(* IEC 61131-3 sources: plc-vscode/tests/st/test-ready/trust-platform/examples/OSCAT/warehouse_conveyor_merge_mediator/oop/src, 3 files *)

(* ---- Main.st ---- *)
(* Pattern role: IInfeedConveyor is the contract boundary for the Mediator example. *)
INTERFACE IInfeedConveyor
    PROPERTY LaneId : INT
    GET
    END_GET
    END_PROPERTY
    PROPERTY Requesting : BOOL
    GET
    END_GET
    END_PROPERTY
    PROPERTY Jammed : BOOL
    GET
    END_GET
    END_PROPERTY
    PROPERTY Granted : BOOL
    GET
    END_GET
    END_PROPERTY
    METHOD UpdateLane
    VAR_INPUT
        Request : BOOL;
        Jam : BOOL;
    END_VAR
    END_METHOD
    METHOD Grant
    VAR_INPUT
        Enable : BOOL;
    END_VAR
    END_METHOD
END_INTERFACE

(* Pattern role: InfeedConveyor is a concrete implementation in the Mediator example. *)
FUNCTION_BLOCK InfeedConveyor IMPLEMENTS IInfeedConveyor
VAR
    LaneIdValue : INT;
    RequestingValue : BOOL;
    JammedValue : BOOL;
    GrantedValue : BOOL;
END_VAR
METHOD PUBLIC Configure
VAR_INPUT
    LaneId : INT;
END_VAR
LaneIdValue := LaneId;
END_METHOD
METHOD PUBLIC UpdateLane
VAR_INPUT
    Request : BOOL;
    Jam : BOOL;
END_VAR
RequestingValue := Request;
JammedValue := Jam;
END_METHOD
METHOD PUBLIC Grant
VAR_INPUT
    Enable : BOOL;
END_VAR
GrantedValue := Enable;
END_METHOD
PUBLIC PROPERTY LaneId : INT
GET
    LaneId := LaneIdValue;
END_GET
END_PROPERTY
PUBLIC PROPERTY Requesting : BOOL
GET
    Requesting := RequestingValue;
END_GET
END_PROPERTY
PUBLIC PROPERTY Jammed : BOOL
GET
    Jammed := JammedValue;
END_GET
END_PROPERTY
PUBLIC PROPERTY Granted : BOOL
GET
    Granted := GrantedValue;
END_GET
END_PROPERTY
END_FUNCTION_BLOCK

(* Composition role: MergeMediator owns the collaborating objects used by this Mediator example. *)
FUNCTION_BLOCK MergeMediator
VAR
    Lane1 : InfeedConveyor;
    Lane2 : InfeedConveyor;
    Lane3 : InfeedConveyor;
    ActiveLaneIdValue : INT;
    GrantedCounter : DwordCounter;
    JamCountValue : INT;
END_VAR
METHOD PUBLIC Initialize
Lane1.Configure(LaneId := INT#1);
Lane2.Configure(LaneId := INT#2);
Lane3.Configure(LaneId := INT#3);
GrantedCounter.Initialize();
GrantedCounter.Configure(StepSize := DWORD#1, MaxValue := DWORD#16#FFFFFFFF);
END_METHOD
METHOD PRIVATE TryGrant : BOOL
VAR_INPUT
    Lane : IInfeedConveyor;
    DownstreamReady : BOOL;
END_VAR
IF (ActiveLaneIdValue = INT#0) AND DownstreamReady AND Lane.Requesting AND NOT Lane.Jammed THEN
    ActiveLaneIdValue := Lane.LaneId;
    Lane.Grant(Enable := TRUE);
    GrantedCounter.Update(Up := TRUE, Down := FALSE);
    TryGrant := TRUE;
ELSE
    Lane.Grant(Enable := FALSE);
    TryGrant := FALSE;
END_IF;
IF Lane.Jammed THEN
    JamCountValue := JamCountValue + INT#1;
END_IF;
END_METHOD
METHOD PUBLIC Update : INT
VAR_INPUT
    Lane1Request : BOOL;
    Lane1Jam : BOOL;
    Lane2Request : BOOL;
    Lane2Jam : BOOL;
    Lane3Request : BOOL;
    Lane3Jam : BOOL;
    DownstreamReady : BOOL;
END_VAR
ActiveLaneIdValue := INT#0;
JamCountValue := INT#0;
(* DwordCounter wraps COUNT_DR (edge-triggered: UP AND NOT LastUp).
   Drop the UP edge first so consecutive scans with grants each emit
   a fresh rising edge and actually increment GrantedCount. *)
GrantedCounter.Update(Up := FALSE, Down := FALSE);
Lane1.UpdateLane(Request := Lane1Request, Jam := Lane1Jam);
Lane2.UpdateLane(Request := Lane2Request, Jam := Lane2Jam);
Lane3.UpdateLane(Request := Lane3Request, Jam := Lane3Jam);
TryGrant(Lane := Lane2, DownstreamReady := DownstreamReady);
TryGrant(Lane := Lane1, DownstreamReady := DownstreamReady);
TryGrant(Lane := Lane3, DownstreamReady := DownstreamReady);
Update := ActiveLaneIdValue;
END_METHOD
PUBLIC PROPERTY ActiveLaneId : INT
GET
    ActiveLaneId := ActiveLaneIdValue;
END_GET
END_PROPERTY
PUBLIC PROPERTY GrantedCount : DWORD
GET
    GrantedCount := GrantedCounter.Count;
END_GET
END_PROPERTY
PUBLIC PROPERTY JamCount : INT
GET
    JamCount := JamCountValue;
END_GET
END_PROPERTY
END_FUNCTION_BLOCK

(* Scan role: Main wires the example objects and exposes the PLC call path under test. *)
PROGRAM Main
VAR
    Merge : MergeMediator;
    Lane1Request : BOOL;
    Lane2Request : BOOL;
    Lane3Request : BOOL;
    DownstreamReady : BOOL;
    Lane1GrantOut : BOOL;
    Lane2GrantOut : BOOL;
    Lane3GrantOut : BOOL;
END_VAR
Merge.Initialize();
Merge.Update(Lane1Request := Lane1Request, Lane1Jam := FALSE, Lane2Request := Lane2Request, Lane2Jam := FALSE, Lane3Request := Lane3Request, Lane3Jam := FALSE, DownstreamReady := DownstreamReady);
Lane1GrantOut := Merge.ActiveLaneId = INT#1;
Lane2GrantOut := Merge.ActiveLaneId = INT#2;
Lane3GrantOut := Merge.ActiveLaneId = INT#3;
END_PROGRAM

(* ---- Configuration.st ---- *)
CONFIGURATION WarehouseConveyorMergeMediatorOopConfiguration
RESOURCE Cpu0 ON PLC
    TASK MainTask (INTERVAL := T#50ms, PRIORITY := 1);
    PROGRAM Merge WITH MainTask : Main;
END_RESOURCE
VAR_CONFIG
    Merge.Lane1Request AT %IX0.0 : BOOL;
    Merge.Lane2Request AT %IX0.1 : BOOL;
    Merge.Lane3Request AT %IX0.2 : BOOL;
    Merge.DownstreamReady AT %IX0.3 : BOOL;
    Merge.Lane1GrantOut AT %QX0.0 : BOOL;
    Merge.Lane2GrantOut AT %QX0.1 : BOOL;
    Merge.Lane3GrantOut AT %QX0.2 : BOOL;
END_VAR
END_CONFIGURATION

(* ---- Tests.st ---- *)
TEST_PROGRAM MergeMediatorGrantsPriorityLane
VAR
    Merge : MergeMediator;
END_VAR
Merge.Initialize();
ASSERT_EQUAL(EXPECTED := INT#2, ACTUAL := Merge.Update(Lane1Request := TRUE, Lane1Jam := FALSE, Lane2Request := TRUE, Lane2Jam := FALSE, Lane3Request := TRUE, Lane3Jam := FALSE, DownstreamReady := TRUE));
ASSERT_EQUAL(EXPECTED := DWORD#1, ACTUAL := Merge.GrantedCount);
END_TEST_PROGRAM

TEST_PROGRAM MergeMediatorSkipsJammedLane
VAR
    Merge : MergeMediator;
END_VAR
Merge.Initialize();
ASSERT_EQUAL(EXPECTED := INT#1, ACTUAL := Merge.Update(Lane1Request := TRUE, Lane1Jam := FALSE, Lane2Request := TRUE, Lane2Jam := TRUE, Lane3Request := FALSE, Lane3Jam := FALSE, DownstreamReady := TRUE));
ASSERT_EQUAL(EXPECTED := INT#1, ACTUAL := Merge.JamCount);
END_TEST_PROGRAM

(* Multi-cycle mediator test: drives the same merge through varying
   lane requests and downstream-ready states. Catches bugs where
   GrantedCount fails to grow on subsequent grants or where the
   mediator gates on stale downstream-ready. *)
TEST_PROGRAM MergeMediatorAccumulatesGrantsAcrossScans
VAR
    Merge : MergeMediator;
END_VAR
Merge.Initialize();

(* Scan 1: lane 2 wins *)
Merge.Update(Lane1Request := TRUE, Lane1Jam := FALSE, Lane2Request := TRUE, Lane2Jam := FALSE, Lane3Request := TRUE, Lane3Jam := FALSE, DownstreamReady := TRUE);
ASSERT_EQUAL(EXPECTED := DWORD#1, ACTUAL := Merge.GrantedCount);

(* Scan 2: only lane 1 requesting, lane 1 grants *)
Merge.Update(Lane1Request := TRUE, Lane1Jam := FALSE, Lane2Request := FALSE, Lane2Jam := FALSE, Lane3Request := FALSE, Lane3Jam := FALSE, DownstreamReady := TRUE);
ASSERT_EQUAL(EXPECTED := DWORD#2, ACTUAL := Merge.GrantedCount);

(* Scan 3: downstream not ready, no grant even with requests *)
Merge.Update(Lane1Request := TRUE, Lane1Jam := FALSE, Lane2Request := TRUE, Lane2Jam := FALSE, Lane3Request := TRUE, Lane3Jam := FALSE, DownstreamReady := FALSE);
ASSERT_EQUAL(EXPECTED := DWORD#2, ACTUAL := Merge.GrantedCount);
END_TEST_PROGRAM

(* Multi-call regression: a long burst of grants accumulates one
   GrantedCount per scan when downstream stays ready. Catches edge-
   trigger bugs in the embedded DwordCounter where a missing edge
   reset would freeze the counter at 1. *)
TEST_PROGRAM MergeMediatorIncrementsCounterOncePerGrantedScan
VAR
    Merge : MergeMediator;
    I : INT;
END_VAR
Merge.Initialize();
FOR I := 1 TO 10 DO
    Merge.Update(Lane1Request := FALSE, Lane1Jam := FALSE, Lane2Request := TRUE, Lane2Jam := FALSE, Lane3Request := FALSE, Lane3Jam := FALSE, DownstreamReady := TRUE);
END_FOR;
ASSERT_EQUAL(EXPECTED := DWORD#10, ACTUAL := Merge.GrantedCount);
END_TEST_PROGRAM

(* Boundary test: no requests at all returns ActiveLaneId = 0 and
   does not increment GrantedCount. *)
TEST_PROGRAM MergeMediatorNoRequestsReturnsZero
VAR
    Merge : MergeMediator;
END_VAR
Merge.Initialize();
ASSERT_EQUAL(EXPECTED := INT#0, ACTUAL := Merge.Update(Lane1Request := FALSE, Lane1Jam := FALSE, Lane2Request := FALSE, Lane2Jam := FALSE, Lane3Request := FALSE, Lane3Jam := FALSE, DownstreamReady := TRUE));
ASSERT_EQUAL(EXPECTED := DWORD#0, ACTUAL := Merge.GrantedCount);
END_TEST_PROGRAM

(* Boundary test: all three lanes jammed. JamCount = 3, ActiveLaneId
   stays 0, GrantedCount unchanged. *)
TEST_PROGRAM MergeMediatorAllLanesJammedNoGrant
VAR
    Merge : MergeMediator;
END_VAR
Merge.Initialize();
ASSERT_EQUAL(EXPECTED := INT#0, ACTUAL := Merge.Update(Lane1Request := TRUE, Lane1Jam := TRUE, Lane2Request := TRUE, Lane2Jam := TRUE, Lane3Request := TRUE, Lane3Jam := TRUE, DownstreamReady := TRUE));
ASSERT_EQUAL(EXPECTED := INT#3, ACTUAL := Merge.JamCount);
ASSERT_EQUAL(EXPECTED := DWORD#0, ACTUAL := Merge.GrantedCount);
END_TEST_PROGRAM

(* Per-FB isolation: drive a bare InfeedConveyor and verify its
   property surface. Each lane object should keep its own jam,
   request, and grant state without depending on a mediator. *)
TEST_PROGRAM InfeedConveyorReportsItsOwnState
VAR
    Lane : InfeedConveyor;
END_VAR

Lane.Configure(LaneId := INT#7);
ASSERT_EQUAL(EXPECTED := INT#7, ACTUAL := Lane.LaneId);
ASSERT_FALSE(IN := Lane.Requesting);
ASSERT_FALSE(IN := Lane.Jammed);
ASSERT_FALSE(IN := Lane.Granted);

Lane.UpdateLane(Request := TRUE, Jam := FALSE);
ASSERT_TRUE(IN := Lane.Requesting);
ASSERT_FALSE(IN := Lane.Jammed);

Lane.Grant(Enable := TRUE);
ASSERT_TRUE(IN := Lane.Granted);

Lane.UpdateLane(Request := TRUE, Jam := TRUE);
ASSERT_TRUE(IN := Lane.Jammed);
END_TEST_PROGRAM

(* Edge input: lane 2 requesting but jammed, lane 3 requesting and
   healthy — lane 3 wins because lane 2 is skipped and lane 1 is not
   requesting. *)
TEST_PROGRAM MergeMediatorJammedHighPriorityFallsThroughToLowestLane
VAR
    Merge : MergeMediator;
END_VAR
Merge.Initialize();
ASSERT_EQUAL(EXPECTED := INT#3, ACTUAL := Merge.Update(Lane1Request := FALSE, Lane1Jam := FALSE, Lane2Request := TRUE, Lane2Jam := TRUE, Lane3Request := TRUE, Lane3Jam := FALSE, DownstreamReady := TRUE));
ASSERT_EQUAL(EXPECTED := INT#1, ACTUAL := Merge.JamCount);
END_TEST_PROGRAM
